Fanuc KAREL source: KT00494.KL

PROGRAM KT00494
%NOLOCKGROUP
VAR
  P1: XYZWPR
  P2: POSITION
  OUT: POSITION
BEGIN
  P1.X = 1.0
  OUT = P1 : P2
END KT00494
